// Generated by voz_llm_plc_agent
// Target: Siemens TIA Portal V18 - SCL external source
// Review and compile before any download to physical hardware.

FUNCTION_BLOCK "PLC_PRG"
{ S7_Optimized_Access := 'TRUE' }
VERSION : 0.1
VAR_INPUT
   I_Emergency : Bool := FALSE;
   I_Fault : Bool := FALSE;
   I_Run_State : Bool := FALSE;
END_VAR
VAR_OUTPUT
   Q_Motor_Enable : Bool := FALSE;
   Q_Alarm : Bool := FALSE;
   Q_Pilot_Run : Bool := FALSE;
   Q_Pilot_Fault : Bool := FALSE;
   Q_Pilot_Stop : Bool := FALSE;
END_VAR
BEGIN
(* Pilotos de estado: falla, marcha o detenido; solo uno encendido (la falla tiene prioridad) *)
#Q_Pilot_Fault := #I_Fault OR #I_Emergency;
#Q_Pilot_Run := #I_Run_State AND NOT #Q_Pilot_Fault;
#Q_Pilot_Stop := NOT #I_Run_State AND NOT #Q_Pilot_Fault;
END_FUNCTION_BLOCK

DATA_BLOCK "DB_PLC_PRG"
{ S7_Optimized_Access := 'TRUE' }
VERSION : 0.1
NON_RETAIN
"PLC_PRG"
BEGIN
END_DATA_BLOCK

ORGANIZATION_BLOCK "Main"
{ S7_Optimized_Access := 'TRUE' }
VERSION : 0.1
BEGIN
   "DB_PLC_PRG"(
      I_Emergency := "I_Emergency",
      Q_Motor_Enable => "Q_Motor_Enable",
      Q_Alarm => "Q_Alarm",
      Q_Pilot_Run => "Q_Pilot_Run",
      Q_Pilot_Fault => "Q_Pilot_Fault",
      I_Fault := "I_Fault",
      I_Run_State := "I_Run_State",
      Q_Pilot_Stop => "Q_Pilot_Stop"
   );
END_ORGANIZATION_BLOCK
